Fanuc KAREL source: kt00216.KL

PROGRAM KT00216
%STACKSIZE=65535
%PRIORITY=65535
%NOLOCKGROUP
VAR
Y1 : ARRAY[2] OF BYTE
H2 : ARRAY[2] OF SHORT
OUT : INTEGER
BEGIN
Y1[1]=2
H2[1]=3
-- UNRESOLVED_PC line 10 opcodes [22 9D 33 B1 22 9D 33 B3 46 23] marker_code=38
END KT00216
